(* IEC 61131-3 sources: plcassist-cli/packages/volt-lsp-iec/test-corpus/awa-palletizer/Device/Plc Logic/Application/Library Manager/L_TS2P_TechModulesSynchronizingCamming (part 3) *)

(* ---- L_TS2P_TM_SYNCPOSBASE.fb ---- *)
FUNCTION_BLOCK L_TS2P_TM_SYNCPOSBASE EXTENDS L_TB2M_TM_MotionControl
VAR
	TM_SYNCPOS : L_TB2P_ModuleHandlerConfig;
	ITFSYNCPOSBASE : L_TS2P_ISyncPosBase := THIS^;
	SCDATA_INT : L_TS2P_scData_TM_SyncPosBase;
	_ITFSTRUCTPROVIDERSYNCPOS : L_TS2P_IStructProviderSyncPos;
	PDATA : POINTER TO L_TS2P_scData_TM_SyncPosBase := ADR(scData_Int);
	PPAR : POINTER TO L_TS2P_scPar_TM_SyncPosBase;
	PSF : POINTER TO L_TS2P_scSF_TM_SyncPosBase;
	PAP : POINTER TO L_TS2P_scAP_TM_SyncPosBase;
	PINPUT2 : POINTER TO L_TS2P_SyncPosBaseIn;
	POUTPUT2 : POINTER TO L_TS2P_SyncPosBaseOut;
	FB_CONDAXISMOVING : L_TB2P_AxisMoving;
	FB_CONDMASTERDIRECTION : L_TB2P_ConditionMasterDirection;
	FB_CONDBASEVELOCITYDIRECTION : L_TB2P_ConditionBaseVelocityDirection;
	FB_CONDSYNCPARAMETER : L_TS2P_ConditionSyncParameter;
	FB_CONDITIONCHECKHOMINGNEEDED : L_UBUP_ConditionInput;
	FB_CONDITIONJOGGINGACTIVE : L_UBUP_ConditionInput;
	FB_CONDCOLLECTSYNCIN : L_UBUP_ConditionCollectionAND := STRUCT(aitfCondition := [fb_ConditionOperationEnabled, fb_ConditionLimiter, fb_CondMasterDirection, fb_CondSyncParameter, fb_ConditionJoggingActive, fb_ConditionAxisNotStopping, fb_ConditionCheckHomingNeeded]);
	FB_CONDCOLLECTBASEVELOCITY : L_UBUP_ConditionCollectionAND := STRUCT(aitfCondition := [fb_CondBaseVelocityDirection, fb_CondCollectOperationEnabledLimiter, fb_ConditionJoggingActive, fb_ConditionAxisNotStopping]);
	FB_TRANSITION2BASEVELOCITYACCDEC : L_UBUP_RequestTransitionLevel;
	FB_TRANSITION2BASEVELOCITY : L_UBUP_RequestTransitionEdge;
	FB_TRANSITION2BASEVELOCITYZERO : L_UBUP_RequestTransitionLevel;
	FB_TRANSITION2SYNCIN : L_UBUP_RequestTransitionLevel;
	FB_TRANSITION2SYNCOUT : L_UBUP_RequestTransitionEdge;
	FB_TRANSITION2SYNCHRONIZED : L_UBUP_RequestTransitionLevel;
	FB_OFFSETANDTRIMX : L_TS2P_OffsetAndTrim;
	FB_ADDOFFSETCYCLICX : L_MC1P_AddOffsetCyclic;
	FB_GEARBOXPOSITION : L_MB1P_GearboxPositionInput;
	FB_AXISCONVERTER : L_MC2P_AxisConverterBase;
	FB_SYNCPOSRESTOREOFFSET : L_TS2P_OffsetAndTrim;
	FB_CLUTCHEXTENDEDBASE : L_TB2P_ClutchExtendedBase;
	FB_ALLOWEDDIRECTION : L_TS2P_AllowedDirection;
	FB_CONTROLSETVALUES : L_MC1P_ControlSetValues;
	MASTERVALUES_INT : L_MC1P_SetAxisRefMasterValues;
	_ITFREQUESTCONDITIONWARNINGHIGHPRIO : L_UBUP_IRequest;
	CONNECTOR : __SYSTEM.IQueryInterface;
	SYNCPOSBASEEXTENSION : L_TS2P_ISyncPosBase;
END_VAR
END_FUNCTION_BLOCK

METHOD HANDLEREJECTEDREQUEST : BOOL
VAR_INPUT
	ITFREQUESTANNOUNCED : L_UBUP_IRequest;
END_VAR
VAR_OUTPUT
	ITFALTERNATIVEREQUEST : L_UBUP_IRequest;
END_VAR
END_METHOD

METHOD CALLFBS
VAR_INPUT
	ECASE : L_UBUP_StateHandleCase;
END_VAR
END_METHOD

METHOD CALLSTATE
VAR_INPUT
	ITFSTATESERVER : L_UBUP_IStateServer;
	ISTATE : INT;
	ECASE : L_UBUP_StateHandleCase;
END_VAR
END_METHOD

METHOD CHECKTRANSITION
VAR_INPUT
	ITFSTATESERVER : L_UBUP_IStateServer;
END_VAR
END_METHOD

METHOD FINALIZECYCLE
END_METHOD

METHOD PREPARECYCLE
END_METHOD

METHOD STIMULATETRANSITION
VAR_INPUT
	ECASE : L_UBUP_StateHandleCase;
END_VAR
END_METHOD

METHOD CALL_SETLOCALMASTERVALUES
END_METHOD

METHOD STATE_01_BASEVEL_ACC_DEC
VAR_INPUT
	ECASE : L_UBUP_StateHandleCase;
	ISTATESERVER : L_UBUP_IStateServer;
END_VAR
END_METHOD

METHOD STATE_02_BASEVEL_2_STANDSTILL
VAR_INPUT
	ECASE : L_UBUP_StateHandleCase;
	ISTATESERVER : L_UBUP_IStateServer;
END_VAR
END_METHOD

METHOD STATE_03_BASEVELOCITY
VAR_INPUT
	ECASE : L_UBUP_StateHandleCase;
	ISTATESERVER : L_UBUP_IStateServer;
END_VAR
END_METHOD

METHOD STATE_11_SYNC_ACC
VAR_INPUT
	ECASE : L_UBUP_StateHandleCase;
	ISTATESERVER : L_UBUP_IStateServer;
END_VAR
END_METHOD

METHOD STATE_12_SYNC_DEC
VAR_INPUT
	ECASE : L_UBUP_StateHandleCase;
	ISTATESERVER : L_UBUP_IStateServer;
END_VAR
END_METHOD

METHOD STATE_13_SYNCHRONISED
VAR_INPUT
	ECASE : L_UBUP_StateHandleCase;
	ISTATESERVER : L_UBUP_IStateServer;
END_VAR
END_METHOD

METHOD ADDOFFSET
VAR_INPUT
	ITFTECHMODULE : L_TS2P_ISyncPosBase;
	LRSETPOS : LREAL;
	LRSETVEL : LREAL;
	LRSETOFFSET : LREAL;
	LRSETOFFSETVEL : LREAL;
	ETRAVERSINGRANGE : L_MC1P.L_MC1P_TraversingRange;
	LRCYCLELENGTH : LREAL;
END_VAR
VAR_OUTPUT
	XERROR : BOOL;
	EERRORID : L_IE1P.L_IE1P_Error;
	LRSETPOSOUT : LREAL;
	LRSETVELOUT : LREAL;
END_VAR
END_METHOD

METHOD CLUTCH
VAR_INPUT
	ITFTECHMODULE : L_TS2P_ISyncPosBase;
	XENABLE : BOOL;
	XSYNCIN : BOOL;
	LRSETBASEVELOCITY : LREAL;
	ESYNCMODE : L_TB2P_SyncMode;
	EALLOWEDDIRECTION : L_TB2P_AllowedDirection;
	LRSYNCVEL : LREAL;
	LRSYNCACC : LREAL;
	LRSYNCDEC : LREAL;
	LRSYNCJERK : LREAL;
	LRSYNCINDIST : LREAL;
	LRSYNCOUTDIST : LREAL;
	LRSYNCOUTPOS : LREAL;
	XLOADCLUTCHOFFSET : BOOL;
	LRLOADCLUTCHOFFSET : LREAL;
	LRCYCLICMASTERPOS : LREAL;
	LRCYCLICMASTERVEL : LREAL;
	ETRAVERSINGRANGEMASTER : L_MC1P_TraversingRange;
	LRCYCLELENGTHMASTER : LREAL;
	LRCYCLICAXISPOS : LREAL;
	LRCYCLICAXISVEL : LREAL;
	LRCYCLICAXISACC : LREAL;
	ETRAVERSINGRANGEAXIS : L_MC1P_TraversingRange;
	LRCYCLELENGTHAXIS : LREAL;
END_VAR
VAR_OUTPUT
	XERROR : BOOL;
	EERRORID : L_IE1P.L_IE1P_Error;
	XBUSY : BOOL;
	XDONE : BOOL;
	XSYNCHRONISED : BOOL;
	XACCDECSYNC : BOOL;
	XINBASEVELOCITY : BOOL;
	LRSETPOSOUT : LREAL;
	LRSETVELOUT : LREAL;
	LRSETACCOUT : LREAL;
	LRCLUTCHOFFSETOUT : LREAL;
END_VAR
END_METHOD

METHOD GEARBOX
VAR_INPUT
	ITFTECHMODULE : L_TS2P_ISyncPosBase;
	XENABLE : BOOL;
	LRSETPOSX : LREAL;
	LRSETVELX : LREAL;
	DWNUMERATOR : DWORD;
	DWDENOMINATOR : DWORD;
	LRCYCLELENGTHX : LREAL;
	LRCYCLELENGTHY : LREAL;
	ETRAVERSINGRANGEX : L_MC1P.L_MC1P_TraversingRange;
	ETRAVERSINGRANGEY : L_MC1P.L_MC1P_TraversingRange;
	XLOADGEARBOXPOS : BOOL;
	LRLOADGEARBOXPOS : LREAL;
END_VAR
VAR_OUTPUT
	XERROR : BOOL;
	EERRORID : L_IE1P.L_IE1P_Error;
	LRSETPOSOUT : LREAL;
	LRSETVELOUT : LREAL;
END_VAR
END_METHOD

METHOD OFFSETANDTRIM
VAR_INPUT
	ITFTECHMODULE : L_TS2P_ISyncPosBase;
	XENABLE : BOOL;
	LRSETOFFSET : LREAL;
	XTRIMPOS : BOOL;
	XTRIMNEG : BOOL;
	LRSETTRIMDISTANCE : LREAL;
	ETRIMMODE : L_TS2P_TrimMode;
	XLOADOFFSET : BOOL;
	XRESETTRIMOFFSET : BOOL;
	LRSETVEL : LREAL;
	LRSETACC : LREAL;
	LRSETDEC : LREAL;
	LRSETJERK : LREAL;
	WACTDIRECTION : WORD;
	EALLOWEDDIRECTION : L_TB2P.L_TB2P_AllowedDirection;
	LRCYCMASTERPOS : LREAL;
	LRCYCMASTERVEL : LREAL;
	LRCYCMASTERACC : LREAL;
END_VAR
VAR_OUTPUT
	XERROR : BOOL;
	EERRORID : L_IE1P.L_IE1P_Error;
	XBUSY : BOOL;
	XDONE : BOOL;
	LRSETOFFSETOUTTOTAL : LREAL;
	LRSETOFFSETOUTTOTALVEL : LREAL;
	LRSETOFFSETOUT : LREAL;
	LRSETOFFSETOUTTRIM : LREAL;
END_VAR
END_METHOD

METHOD CALL_ALLOCPOINTADR
END_METHOD

METHOD CALL_EXIT_CALLFBS
END_METHOD

METHOD CALL_INIT_CALLFBS
END_METHOD

METHOD CALL_RESETOUTPUT
END_METHOD

METHOD MAPTMSTATE
VAR_INPUT
	ETMSTATEINTERNAL : L_TB2P_States;
END_VAR
VAR_OUTPUT
	ETMSTATEEXTERNAL : L_TB2P_States;
END_VAR
END_METHOD

(* ---- L_TS2P_TOOLCORRECTION.fb ---- *)
FUNCTION_BLOCK L_TS2P_TOOLCORRECTION
VAR_INPUT
	XENABLE : BOOL;
	XACTIVATECORRECTION : BOOL;
	TPRECDATA : L_MC1P_TpReceiveData;
	LRSENSORTOOLDISTANCE : LREAL;
	LRMAXCORRNEG : LREAL;
	LRMAXCORRPOS : LREAL;
	LRUPPERCORRPOS : LREAL;
	LRLOWERCORRPOS : LREAL;
	DNNUMAXISY : DWORD;
	DNDENAXISY : DWORD;
	XENABLEMARKWINDOW : BOOL;
	XTEACHMARKWINDOW : BOOL;
	LRMARKWINDOWSIZE : LREAL;
	LRSETOFFSETMARKWINDOW : LREAL;
	DWMAXNUMBERVIRTUALMARKS : DWORD;
	ECORRMODE : L_TS2P_CorrectionMode;
	LRCORRVEL : LREAL;
	LRCORRACC : LREAL;
	LRCORRDEC : LREAL;
	LRCORRJERK : LREAL;
END_VAR
VAR_OUTPUT
	XERROR : BOOL;
	XWARNING : BOOL;
	EERRORID : WORD;
	XCORRLIMITED : BOOL;
	LRACTMARKERROR : LREAL;
	LRACTMARKDIST : LREAL;
	XINITDONE : BOOL;
	XCORRACTIVE : BOOL;
	XMARKRECEIVED : BOOL;
	LRSENSORACTPOS : LREAL;
	LRSENSORSETPOS : LREAL;
	XMARKWINDOWOPEN : BOOL;
	XMARKOUTOFWINDOW : BOOL;
	XMARKNOTDETECTED : BOOL;
	XMARKWINDOWTEACHED : BOOL;
END_VAR
VAR_IN_OUT
	AXIS : AXIS_REF;
END_VAR
VAR
	SPEEDTOPOSINTEGRATE : L_MC1P_IntegrateAxis;
	TPLIMITDIFF : L_TS2P_TpLimitDiff;
	FB_ADDOFFSET : L_MC1P_AddOffsetCyclic;
	TPCALCDIFF : L_MC1P_TpCalcDiff;
	TP_CONVERTER : L_TB2P_TP_Converter;
	DISTCORRECTIONWINDOW : L_TS2P_DistCorrectionWindow;
	MARKWINDOW : L_TS2P_MarkWindowRelative;
	MARKSTACK : L_TS2P_MarkStack;
	TPVIRTUALACTPOS : L_TS2P_TpVirtualActPos;
	FB_PROFILEGENERATOR : L_MC1P_ProfileGenerator;
	FB_INTEGRATOR : L_MC1P_IntegrateAxis;
	SCPROFILEPARAMETER : L_MC1P_ProfileParameter;
	LRMARKSENSORPOS : LREAL;
	LRGEARINGFAKTOR : LREAL := 1.0;
	XERROR_TM : BOOL;
	EERRORID_TM : L_IE1P_Error;
	LRTPDIFFERENCE : LREAL;
	XLOADMARKSENSORPOS_OLD : BOOL;
	XTPRECEIVED_OLD : BOOL;
	LRMARKWINDOWSIZE_INT : LREAL;
	XTPINWINDOW : BOOL;
	LRPOS_INT : LREAL;
	XTPRECEIVEDOUT_INT : BOOL;
	LRTPACTPOSITION_INT : LREAL;
	LRTPDIFFERENCELIM_INT : LREAL;
	LROFFSETPOSCTRL_INT : LREAL;
	LRPOSOUT_INT : LREAL;
	LRVELOUT_INT : LREAL;
	XCORRACTIVE_INT : BOOL;
	XINIT : BOOL := TRUE;
	XTPCORRECTIONACTIVE : BOOL := FALSE;
	LRTPAXISSETPOS : LREAL;
	LRMARKDIST_INT : LREAL;
	XZERO : BOOL;
	XHOMINGDONE : BOOL;
	XSTARTREFERENCEACTIVE : BOOL;
	XHOMINGACTIVE : BOOL := FALSE;
	XMARKDISTCHANGED : BOOL;
	LRTPACTPOSIN_OLD : LREAL;
	LRTPAXISACTPOS_OLD : LREAL;
	ICOUNTER : INT := 0;
	XFIRSTTOUCHPROBE : BOOL := TRUE;
	LRMARKSTACKLENGTH : LREAL;
	LRTPDIFFERENCELIMITOUT_INT : LREAL;
	XTPRECEIVESTACKOUT_INT : BOOL;
	XTPNOTDETECTED_INT : BOOL;
	XMAXTPNOTDETECTED : BOOL;
	LRGEARFACTORINTEGRATOR : LREAL;
	LRGEARFACTORGAIN : LREAL := 1;
	LRGEARFACTORNUMERATORCORR : LREAL;
	LRGEARFACTORNUMERATORCORRLIMITED : LREAL;
	LRGEARFACTORDENOMINATOR : LREAL;
	LRGEARFACTORNUMERATOR : LREAL;
	LRTOTALSTACKDIFFERENCEOUT_INT : LREAL := 0;
	LCORRECTIONVELIN : LREAL;
	LRSETPOSCORROUT_OLD : LREAL;
	LRDELTAGEARFACTORCORR : LREAL;
	XTPSENSORTEACHEDOLD : BOOL;
	XTPSENSORTEACHEDATLASTMARK : BOOL;
	XCALCMARKDISTINITIALISED : BOOL;
	XTEACHTPSENSOROLD : BOOL;
	LRTPDEADTIMEDIFF : LREAL;
	XTPRECEIVEDOUTOLD_INT : BOOL;
	LRMARKDISTINTEGRATOR : LREAL;
	LRPOSOUTOLD_INT : LREAL;
	LRCORRPOS_INT : LREAL;
	LRCORRPOSOLD_INT : LREAL := 0;
	XENABLEOLD : BOOL;
	TPRECDATAMARKSTACK : L_MC1P_TpReceiveData;
	TPRECDATAMARKWINDOW : L_MC1P_TpReceiveData;
	XTPRECEIVEDINOLD_INT : BOOL;
	XFIRSTVALUESTORED : BOOL;
	LRAXISSETPOSOLD_INT : LREAL;
	LRCORRRESIDUAL : LREAL;
	ECORRECTIONMODEOLD : L_TS2P_CorrectionMode;
	XCORRECTIONBUSY : BOOL;
END_VAR
END_FUNCTION_BLOCK

METHOD CALL_CALCACTMARKDIST
END_METHOD

METHOD CALL_CALCTOOLERROR
END_METHOD

METHOD CALL_CORRECTIONPOS
END_METHOD

METHOD CALL_CORRECTIONPROFILE
END_METHOD

METHOD CALL_ENABLEREGISTERCONTROL
END_METHOD

METHOD CALL_ERRORHANDLER
END_METHOD

METHOD CALL_FB
END_METHOD

METHOD CALL_INPUT
END_METHOD

METHOD CALL_LIMIT
END_METHOD

METHOD CALL_MARKDISTCHANGE
END_METHOD

METHOD CALL_MARKSENSORPOS
END_METHOD

METHOD CALL_MARKSTACK
END_METHOD

METHOD CALL_MARKWINDOW
END_METHOD

METHOD CALL_NOTENABLE
END_METHOD

METHOD CALL_OUTPUT
END_METHOD

METHOD CALL_RESET
END_METHOD

METHOD CALL_RESETOUTPUTS
END_METHOD

METHOD CALL_SETCORRECTION
END_METHOD

METHOD CALL_TPCONVERTER
END_METHOD

METHOD CALL_VIRTUALACTPOS
END_METHOD

METHOD GET_ACTMARKERRORLIMITED : LREAL
END_METHOD

METHOD GET_ACTUALMARKDIST : LREAL
END_METHOD

METHOD GET_CORRREGPOS : LREAL
END_METHOD

METHOD GET_INTEGRATORREGPOS : LREAL
END_METHOD

METHOD GET_MARKERRORUNLIMITED : LREAL
END_METHOD

METHOD GET_MARKPOSITIONINREGISTER : LREAL
END_METHOD

METHOD GET_MARKRECEIVEUNLIMITED : BOOL
END_METHOD

METHOD GET_MARKRECEIVEDLIMITED : BOOL
END_METHOD

METHOD GET_MARKWINDOWCOMP : BOOL
END_METHOD

METHOD GET_REGISTERINPUTVEL : LREAL
END_METHOD

METHOD GET_SETVELOCITYREGISTER : LREAL
END_METHOD

METHOD GET_LRMARKSTACKLENGTH : LREAL
END_METHOD

(* ---- L_TS2P_TPLIMITDIFF.fb ---- *)
FUNCTION_BLOCK L_TS2P_TPLIMITDIFF
VAR_INPUT
	XENABLE : BOOL;
	XTPRECEIVED : BOOL;
	LRSETTPDIFFERENCE : LREAL;
	LRSETLIMITMIN : LREAL := -100;
	LRSETLIMITMAX : LREAL := 100;
END_VAR
VAR_OUTPUT
	XTPRECEIVEDOUT : BOOL;
	XLIMITACTIVE : BOOL;
	LRTPDIFFERENCELIM : LREAL;
END_VAR
VAR
	XTPRECEIVEDOLD : BOOL;
END_VAR
END_FUNCTION_BLOCK

(* ---- L_TS2P_TPVIRTUALACTPOS.fb ---- *)
FUNCTION_BLOCK L_TS2P_TPVIRTUALACTPOS
VAR_INPUT
	XTPWINDOWOPEN : BOOL;
	XTPRECEIVEDIN : BOOL;
	XMAXTPNOTDETECTED : BOOL;
	LRSETTPPOSIN : LREAL;
	LRACTTPPOSIN : LREAL;
END_VAR
VAR_OUTPUT
	XTPRECEIVEDOUT : BOOL;
	LRACTTPPOS : LREAL;
END_VAR
VAR
	XTPRECEIVEDINOLD : BOOL;
	XFLAGWINDOWOPENANDNOTP : BOOL := FALSE;
	XWINDOWOPENOLD : BOOL;
	XVIRTUALTPACTIVE : BOOL;
END_VAR
END_FUNCTION_BLOCK

(* ---- L_TS2P_VISUPOOL.fb ---- *)
FUNCTION_BLOCK L_TS2P_VISUPOOL
VAR
	M_STNAMESPACE : STRING(80);
	M_STHELPVARID : STRING;
	M_STHELPVARPATH : STRING(255);
	M_STHELP : STRING;
	M_REGISTERIMAGES : BOOL := TRUE;
END_VAR
END_FUNCTION_BLOCK

METHOD FB_INIT : BOOL
VAR_INPUT
	BINITRETAINS : BOOL;
	BINCOPYCODE : BOOL;
END_VAR
END_METHOD

METHOD FB_REINIT : BOOL
END_METHOD

METHOD FB_EXIT : BOOL
VAR_INPUT
	BINCOPYCODE : BOOL;
END_VAR
END_METHOD

(* ---- L_TT1P_INPOSITION.fb ---- *)
FUNCTION_BLOCK L_TT1P_INPOSITION
VAR_INPUT
	XENABLE : BOOL;
	LRPOSWINDOW : LREAL;
	LRPOSTIME : LREAL;
	XHOLDSETPOS : BOOL;
END_VAR
VAR_OUTPUT
	XINPOSITION : BOOL;
	XBUSY : BOOL;
	LRHOLDPOSITION : LREAL;
	XERROR : BOOL;
	EERRORID : L_IE1P_Error;
END_VAR
VAR_IN_OUT
	AXIS : AXIS_REF;
END_VAR
VAR
	XINTOL : BOOL;
	XENABLEOLD : BOOL := FALSE;
	XHOLDSETPOSOLD : BOOL := FALSE;
	LRSETPOSITIONOLD : LREAL;
	XSETPOSITIONCHG : BOOL;
	INPOSITION_TON : TON;
	INPOSITION_F_TRIG : F_TRIG;
	TIMEOUT_TON : TON;
END_VAR
END_FUNCTION_BLOCK

METHOD FB_RESET : BOOL
END_METHOD

(* ---- LOCKTOMASTER.fb ---- *)
FUNCTION_BLOCK LOCKTOMASTER
VAR_INPUT
	XENABLE : BOOL;
	XLOCKTOMASTER : BOOL;
	XRESETOFFSETLOCKTOMASTER : BOOL;
	ELOCKTOMASTERMODE : L_TS2P_SyncInMode;
	EDIRECTION : MC_DIRECTION := 3;
	LRSETPOSIN : LREAL;
	LRSETVELIN : LREAL;
	LRSETACCIN : LREAL;
	LRSETVEL : LREAL := 360.0;
	LRSETACC : LREAL := 3600.0;
	LRSETDEC : LREAL := 3600.0;
	LRSETJERK : LREAL := 10000.0;
	LRPARKPOSITION : LREAL := 0;
	LRCYCLICAXISPOS : LREAL;
	LRCYCLICAXISVEL : LREAL;
	LRCYCLICAXISACC : LREAL;
END_VAR
VAR_OUTPUT
	XERROR : BOOL;
	EERRORID : L_IE1P_Error;
	XLOCKTOMASTERBUSY : BOOL;
	XMASTERLOCKED : BOOL;
	LRSETPOSOUT : LREAL;
	LRSETVELOUT : LREAL;
	LRSETACCOUT : LREAL;
	LROFFSETLOCKTOMASTER : LREAL;
END_VAR
VAR_IN_OUT
	AXIS : AXIS_REF;
END_VAR
VAR
	L_MC1P_ADDOFFSETCYCLIC1 : L_MC1P_AddOffsetCyclic;
	L_MC1P_PROFILEGENERATOR1 : L_MC1P_ProfileGenerator;
	XINTOLERANCEWINDOW : BOOL;
	XLOCKTOMASTER_OLD : BOOL;
	EDIRECTION_INT : MC_DIRECTION;
	LRSTARTPOS_INT : LREAL;
	LRSETPOSADDOFFSETCYCLIC : LREAL;
	XRESETACTIVE : BOOL;
	XRESETOFFSETLOCKTOMASTER_OLD : BOOL;
	LRSETOFFSET : LREAL;
	LRSETVELOLD : LREAL;
	LRSETACCOLD : LREAL;
	LRSETJERKOLD : LREAL;
END_VAR
END_FUNCTION_BLOCK

METHOD CALCULATELOCKTOCAMDIRECTION
VAR_INPUT
	LRTARGETPOS : LREAL;
	LRACTUALPOS : LREAL;
	LRACTUALVELOCITY : LREAL;
	EDIRECTION : MC_DIRECTION;
	ETRAVERSINGRANGE : L_MC1P_TraversingRange;
	XINTOLERANCEWINDOW : BOOL;
END_VAR
VAR_OUTPUT
	ECLUTCHDIRECTION : L_MC2P_ClutchDirection;
	LRSTARTPOS : LREAL;
END_VAR
END_METHOD
